(*
SPDX-FileCopyrightText: © 2026 Oleksandr Tiutyk <trofimich@gmail.com>
SPDX-License-Identifier: MIT
License: https://opensource.org/license/mit
*)

(* Selects the OnConfigure behavior executed by StaticConfigurationTestWorkflow. *)

{attribute 'qualified_only'}
{attribute 'strict'}
{attribute 'to_string'}
TYPE STATIC_WORKFLOW_TEST_MODE :
(
	NORMAL := 0,
	THROW_BEFORE_SET_ROOT,
	THROW_AFTER_SET_ROOT,
	REENTER_REQUEST_START,
	REENTER_EXECUTE,
	REENTER_DISPOSE_DYNAMIC_CHILDREN,
	REENTER_REQUEST_SUSPEND,
	REENTER_REQUEST_CANCEL,
	REENTER_REQUEST_RESET
);
END_TYPE

(* stored: Version 1.1.0.1, ProductVersion 3.1.4026.21
   DUT STATIC_WORKFLOW_TEST_MODE: Id {9868e2c9-1f15-4117-860e-e03b275a9d22} *)
